TYPE "FRK_HostBook"
VERSION : 0.1
   STRUCT
      "View" {ExternalAccessible := 'False'; ExternalVisible := 'False'; ExternalWritable := 'False'} : "FRK_HostEvents";
      "Sequence" {ExternalAccessible := 'False'; ExternalVisible := 'False'; ExternalWritable := 'False'} : UDInt;
   END_STRUCT;
END_TYPE
